Fanuc KAREL source: kt00893.KL

-- PROVISIONAL review KL for V770-1; original PC SHA256 f75cd4253c857bdb38dcb00aa0ac663d18c5b84887a575ee0412233110ccfe31
-- Incomplete behavior may be omitted. Consult companion uncertainty JSON. Do not deploy.
PROGRAM KT00893
%NOLOCKGROUP
VAR
  OUT : BOOLEAN
-- UNRESOLVED_DECL P1 type=000101
-- UNRESOLVED_DECL P2 type=000101
BEGIN
  -- UNRESOLVED_PC offsets 5-31; opcodes 27,27,49,7E,AD,27,9D,76,23
  -- UNRESOLVED_PC offsets 36-40; opcodes 7F
END KT00893
